Staubli VAL3: utCommon.pjx

--- utCommon.pjx ---
Parameters version=s8.8.3Cs9_BS1660 stackSize=5000 millimeterUnit=true
Program file=start.pgx
Program file=stop.pgx
Data file=utCommon.dtx

--- utCommon.dtx ---
public bool bDisabled
public string sValue
public string sID
public string sOption{}
public string sItem
public string sPage

--- start.pgx ---
program start()
begin
end

--- stop.pgx ---
program stop()
begin
end
